// TIA Portal project "s16_stl" (V21)

(* hardware
DEVICE "S7-1500/ET200MP station_1"  S7-1500 station
   slot 0: "Rail_0"  Rack  6ES7 590-1***0-0AA0
   slot 1: "S16PLC"  CPU 1511-1 PN  6ES7 511-1AL03-0AB0  V4.1
      slot 3: "CPU display_1"  6ES7591-1AA00-0AA0
      slot 32768: "PROFINET interface_1"  X1
         slot 32769: "Port_1"  X1 P1
         slot 32770: "Port_2"  X1 P2
      slot 34817: "Virtual CP interface port_1"  Virtual CP interface port  Virtual CP interface port FW V4.1
*)

// ===== PLC "S16PLC"  CPU 1511-1 PN =====

VAR_GLOBAL   // PLC tag table "Default tag table"
   "Start" AT %I0.0 : Bool;
   "Stop" AT %I0.1 : Bool;
   "Level" AT %I0.2 : Bool;
   "Rst" AT %I0.3 : Bool;
   "Up" AT %I0.4 : Bool;
   "Down" AT %I0.5 : Bool;
   "SetC" AT %I0.6 : Bool;
   "Sel" AT %IB1 : Byte;
   "Out1" AT %Q0.0 : Bool;
   "Out2" AT %Q0.1 : Bool;
   "Out3" AT %Q0.2 : Bool;
   "Out4" AT %Q0.3 : Bool;
   "Out5" AT %Q0.4 : Bool;
   "Out6" AT %Q0.5 : Bool;
   "Out7" AT %Q0.6 : Bool;
   "Out8" AT %Q0.7 : Bool;
   "RunOn" AT %T7 : Timer;
   "Parts" AT %C3 : Counter;
   "Tag_1" AT %M20.0 : Bool;
   "Tag_2" AT %MW22 : Word;
   "Tag_3" AT %MW24 : Word;
   "Tag_4" AT %MW26 : Word;
   "Tag_5" AT %MD28 : DWord;
   "Tag_6" AT %MW30 : Word;
   "Tag_7" AT %MD44 : DWord;
   "Tag_8" AT %MW48 : Word;
   "Tag_9" AT %M50.0 : Bool;
   "Tag_10" AT %MW52 : Word;
   "Tag_11" AT %MW54 : Word;
   "Tag_12" AT %T1 : Timer;
   "Tag_13" AT %MW60 : Word;
   "Tag_14" AT %MW62 : Word;
   "Tag_15" AT %MW64 : Word;
   "Tag_16" AT %MW66 : Word;
   "Tag_17" AT %MW68 : Word;
   "Tag_18" AT %T2 : Timer;
   "Tag_19" AT %A1.0 : Bool;
   "Tag_20" AT %Z4 : Counter;
   "Tag_21" AT %MW76 : Word;
   "Tag_22" AT %T3 : Timer;
   "Tag_23" AT %MW70 : Word;
   "Tag_24" AT %MW72 : Word;
   "Tag_25" AT %T4 : Timer;
   "Tag_26" AT %Q1.1 : Bool;
   "Tag_27" AT %C2 : Counter;
   "Tag_28" AT %Q1.2 : Bool;
   "Tag_29" AT %MW74 : Word;
   "Tag_30" AT %C5 : Counter;
   "Tag_31" AT %Q1.3 : Bool;
   "Tag_32" AT %T6 : Timer;
   "Tag_33" AT %Q1.4 : Bool;
END_VAR

DATA_BLOCK "LadS5_DB"   // DB2
{ S7_Optimized_Access := 'TRUE' }
VERSION : 0.1
// stored: InstanceOfName LadS5
"LadS5"
BEGIN
END_DATA_BLOCK

DATA_BLOCK "S16Data"   // DB5
{ S7_Optimized_Access := 'FALSE' }
VERSION : 0.1
   VAR
      b0 : Bool;
      b1 : Bool;
      "by" : Byte;
      w : Int;
      d : DInt;
      r : Real;
      s : String[4];
      arr : Array[1..3] of Int;
   END_VAR
BEGIN
END_DATA_BLOCK

FUNCTION_BLOCK "LadS5"   // FB1, LAD
{ S7_Optimized_Access := 'TRUE' }
VERSION : 0.1
   VAR_TEMP   // added for the SCL form of the ladder/FBD networks
      _w1 : Bool;
   END_VAR
BEGIN

REGION Network 1
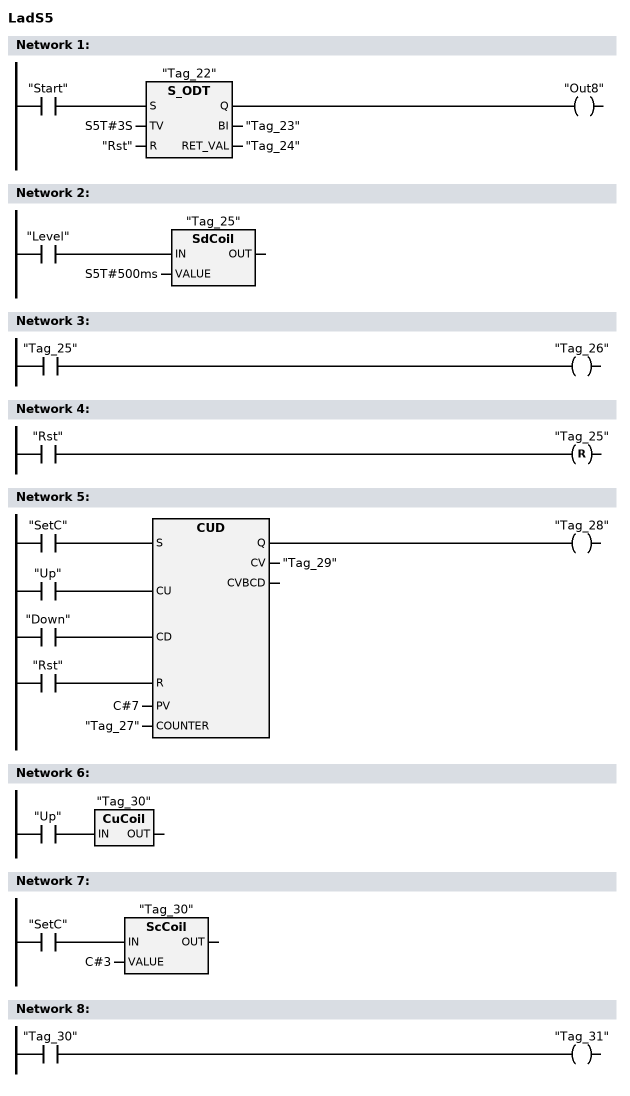
   RUNG wire#powerrail
      Contact( "Start" )
      S_ODT(T_NO := "Tag_22", TV := S5T#3S, R := "Rst", BI => "Tag_23", RET_VAL => "Tag_24")
      Coil( "Out8" )
   END_RUNG
   // the same network as SCL:
   "Tag_24" := S_ODT(T_NO := "Tag_22", S := "Start", TV := S5T#3S, R := "Rst", Q => #_w1, BI => "Tag_23");
   "Out8" := #_w1;
END_REGION

REGION Network 2
   // no SCL statement known for SdCoil: written as a call
   SdCoil(in := "Level", value := S5T#500ms, operand := "Tag_25");
END_REGION

REGION Network 3
   RUNG wire#powerrail
      Contact( "Tag_25" )
      Coil( "Tag_26" )
   END_RUNG
   // the same network as SCL:
   "Tag_26" := "Tag_25";
END_REGION

REGION Network 4
   RUNG wire#powerrail
      Contact( "Rst" )
      R_Coil( "Tag_25" )
   END_RUNG
   // the same network as SCL:
   IF "Rst" THEN "Tag_25" := FALSE; END_IF;
END_REGION

REGION Network 5
   // no SCL statement known for Cud: written as a call
   Cud(cu := "Up",
       cd := "Down",
       s := "SetC",
       r := "Rst",
       pv := C#7,
       "counter" := "Tag_27",
       q => #_w1,
       cv => "Tag_29");
   "Tag_28" := #_w1;
END_REGION

REGION Network 6
   // no SCL statement known for CuCoil: written as a call
   CuCoil(in := "Up", operand := "Tag_30");
END_REGION

REGION Network 7
   // no SCL statement known for ScCoil: written as a call
   ScCoil(in := "SetC", value := C#3, operand := "Tag_30");
END_REGION

REGION Network 8
   RUNG wire#powerrail
      Contact( "Tag_30" )
      Coil( "Tag_31" )
   END_RUNG
   // the same network as SCL:
   "Tag_31" := "Tag_30";
END_REGION
END_FUNCTION_BLOCK

FUNCTION "StlLogic" : Void   // FC1, STL
{ S7_Optimized_Access := 'FALSE' }
VERSION : 0.1
BEGIN

REGION Network 1: AND before OR and a bracket:
         A     "Start";
         A     "Stop";
         O;
         A     "Level";
         AN    "Rst";
         =     "Out1";
         A     "Start";
         O(;
         A     "Level";
         A     "Up";
         );
         =     "Out2";
END_REGION

REGION Network 2: an edge, a jump, a jump list:
         A     "Up";
         FP    "Tag_1";
         JCN   M001;
         L     "Tag_2";
         +     1;
         T     "Tag_2";
   M001: L     "Sel";
         JL    LST;
         JU    L0;
         JU    L1;
   LST:  JU    L2;
   L0:   L     10;
         T     "Tag_3";
         JU    END;
   L1:   L     11;
         T     "Tag_3";
         JU    END;
   L2:   L     12;
         T     "Tag_3";
   END:  NOP   0;
END_REGION

REGION Network 3: arithmetic, a comparison, RND:
         L     "Tag_2";
         L     3;
         *I;
         T     "Tag_4";
         L     "Tag_4";
         L     10;
         >I;
         =     "Out3";
         L     2.5;
         RND;
         T     "Tag_5";
END_REGION
END_FUNCTION

FUNCTION "StlAbs" : Void   // FC2, STL
{ S7_Optimized_Access := 'FALSE' }
VERSION : 0.1
   VAR_TEMP
      "a" : Int;
      "b" : Bool;
      c : Int;
      p : ANY;
      x : Int;
   END_VAR
BEGIN

REGION Network 1: the open DB, absolute and fully qualified:
         OPN   "S16Data";
         SET;
         =     %Data0.1;
         L     7;
         T     %DataB1;
         L     1234;
         T     %DataW2;
         L     "S16Data".w;
         +     1;
         T     "S16Data".arr[1];
         OPN   "S16Data";
         L     2.5;
         T     %DataD8;
         L     DBNO;
         T     "Tag_6";
END_REGION

REGION Network 2: AR1, AR2, register- and memory-indirect:
         OPN   "S16Data";
         L     P#20.0;
         LAR1;
         L     42;
         T     DBW[AR1,P#2.0];
         L     P#M40.0;
         LAR2;
         L     99;
         T     W[AR2,P#0.0];
         L     16;
         T     "Tag_7";
         L     DBW ["Tag_7"];
         T     "Tag_8";
END_REGION

REGION Network 3: local data by address:
         L     5;
         T     #"a";
         L     #"a";
         +     1;
         T     #c;
         SET;
         =     %L2.1;
         A     %L2.1;
         =     "Tag_9";
         L     42;
         T     #x;
         L     #x;
         T     "Tag_10";
         L;
         LAR1;
         L     77;
         T     W[AR1,P#0.0];
         L     #c;
         T     "Tag_11";
END_REGION
END_FUNCTION

FUNCTION "StlS5" : Void   // FC3, STL
{ S7_Optimized_Access := 'FALSE' }
VERSION : 0.1
BEGIN

REGION Network 1: S5 timers, by address and by tag:
         A     "Start";
         L     S5T#2S;
         SD    "Tag_12";
         A     "Tag_12";
         =     "Out4";
         L     "Tag_12";
         T     "Tag_13";
         LC    "Tag_12";
         T     "Tag_14";
         A     "Stop";
         L     S5T#1S;
         SF    "RunOn";
         A     "RunOn";
         =     "Out5";
         A     "Rst";
         R     "Tag_12";
END_REGION

REGION Network 2: an S5 counter by tag:
         A     "Up";
         CU    "Parts";
         A     "Down";
         CD    "Parts";
         A     "SetC";
         L     C#5;
         S     "Parts";
         A     "Rst";
         R     "Parts";
         A     "Parts";
         =     "Out6";
         L     "Parts";
         T     "Tag_15";
         LC    "Parts";
         T     "Tag_16";
END_REGION
END_FUNCTION

FUNCTION "StlGerman" : Void   // FC4, STL
{ S7_Optimized_Access := 'TRUE' }
VERSION : 0.1
BEGIN

REGION Network 1: (SE in German is the on delay; A 1.0 is the output Q1.0)
         A     "Start";
         L     S5T#2S;
         SD    "Tag_18";
         A     "Tag_18";
         =     "Tag_19";
         A     "Level";
         CU    "Tag_20";
         L     "Tag_20";
         T     "Tag_21";
END_REGION
END_FUNCTION

FUNCTION "FbdS5" : Void   // FC5, FBD
{ S7_Optimized_Access := 'TRUE' }
VERSION : 0.1
   VAR_TEMP   // added for the SCL form of the ladder/FBD networks
      _w1 : Bool;
      _s5time1 : S5Time;
   END_VAR
BEGIN

REGION Network 1
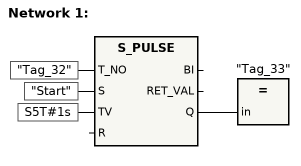
   #_s5time1 := S_PULSE(T_NO := "Tag_32", S := "Start", TV := S5T#1s, Q => #_w1);
   "Tag_33" := #_w1;
END_REGION
END_FUNCTION

ORGANIZATION_BLOCK "Main"   // OB1, LAD, ProgramCycle
TITLE = "Main Program Sweep (Cycle)"
{ S7_Optimized_Access := 'TRUE' }
VERSION : 0.1
   VAR_INPUT
      Initial_Call : Bool;   // Initial call of this OB
      Remanence : Bool;   // =True, if remanent data are available
   END_VAR
BEGIN

REGION Network 1
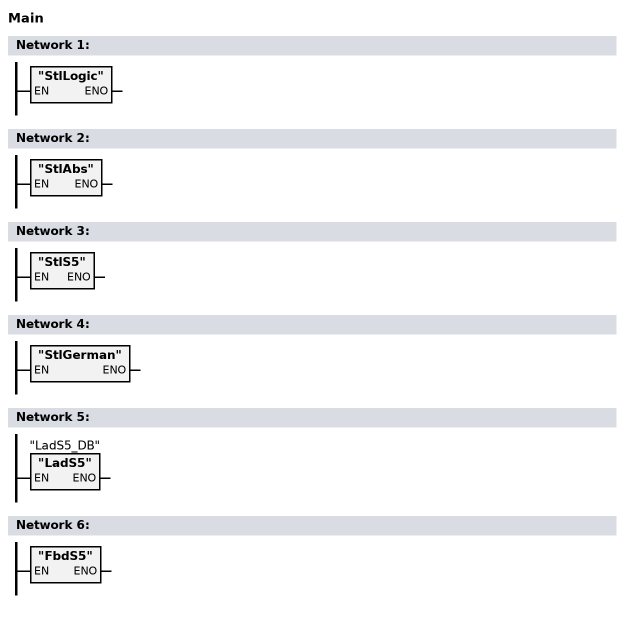
   RUNG wire#powerrail
      "StlLogic"()
   END_RUNG
   // the same network as SCL:
   "StlLogic"();
END_REGION

REGION Network 2
   RUNG wire#powerrail
      "StlAbs"()
   END_RUNG
   // the same network as SCL:
   "StlAbs"();
END_REGION

REGION Network 3
   RUNG wire#powerrail
      "StlS5"()
   END_RUNG
   // the same network as SCL:
   "StlS5"();
END_REGION

REGION Network 4
   RUNG wire#powerrail
      "StlGerman"()
   END_RUNG
   // the same network as SCL:
   "StlGerman"();
END_REGION

REGION Network 5
   RUNG wire#powerrail
      "LadS5_DB"()
   END_RUNG
   // the same network as SCL:
   "LadS5_DB"();   // "LadS5"
END_REGION

REGION Network 6
   RUNG wire#powerrail
      "FbdS5"()
   END_RUNG
   // the same network as SCL:
   "FbdS5"();
END_REGION
END_ORGANIZATION_BLOCK